// TIA Portal V21 export
// export: Created 2026-11-22T02:34:18.9785289Z, ExportSetting WithDefaults, DisplayName Totally Integrated Automation Portal, DisplayVersion V21 Update 3, DisplayName STEP 7 Professional, DisplayVersion V21 Update 3, DisplayName STEP 7 Safety, DisplayVersion V21, DisplayName Tech WebApplication, DisplayVersion V21, DisplayName WinCC Basic/Comfort/Advanced, DisplayVersion V21 Update 3, DisplayName WinCC Unified, DisplayVersion V21 Update 3
Screen "D_Slider_2"  800x480, Number=481
  ScreenLayer "Layer_0"
    Slider "PV_Int" at 6,4 size 60x160  MaximumValue=100, StyleItem=Slider, Caption="SIMATIC"
      ProcessValue := D_Int
    TextField "Label_PV_Int" at 6,196 size 108x16  StyleItem=Text field, Text="PV_Int"
    Slider "PV_Pct_0_200" at 118,4 size 60x160  MaximumValue=200, StyleItem=Slider, Caption="SIMATIC"
      ProcessValue := D_Pct
    TextField "Label_PV_Pct_0_200" at 118,196 size 108x16  StyleItem=Text field, Text="PV_Pct_0_200"
    IOField "State" at 4,454 size 60x22  DataFormat=Decimal, FormatPattern=9, Mode=Output, StyleItem=I/O field
      ProcessValue := D_State
    Button "S1" at 70,454 size 40x22  Mode=Text, StyleItem=Button, TextOff="S1", TextOn="S1"
      on Click: SetS1()
    Button "S2" at 114,454 size 40x22  Mode=Text, StyleItem=Button, TextOff="S2", TextOn="S2"
      on Click: SetS2()
    Button "S3" at 158,454 size 40x22  Mode=Text, StyleItem=Button, TextOff="S3", TextOn="S3"
      on Click: SetS3()
    Button "S4" at 202,454 size 40x22  Mode=Text, StyleItem=Button, TextOff="S4", TextOn="S4"
      on Click: SetS4()
    Button "Next" at 756,454 size 40x22  Mode=Text, StyleItem=Button, TextOff="Next", TextOn="Next"
      on Click: ActivateScreen(Screen name := D_Gauge_1, Object number := 0)
